TYPE "ST_StepTiming"
VERSION : 0.1
   STRUCT
      StepNo : Int;
      StepName : String[120];
      TimeClass : DInt;
      Started : LDT;
      StartedTimeSynchronized : Bool;
      Duration : Time;
      Expected : Time;
   END_STRUCT;

END_TYPE

